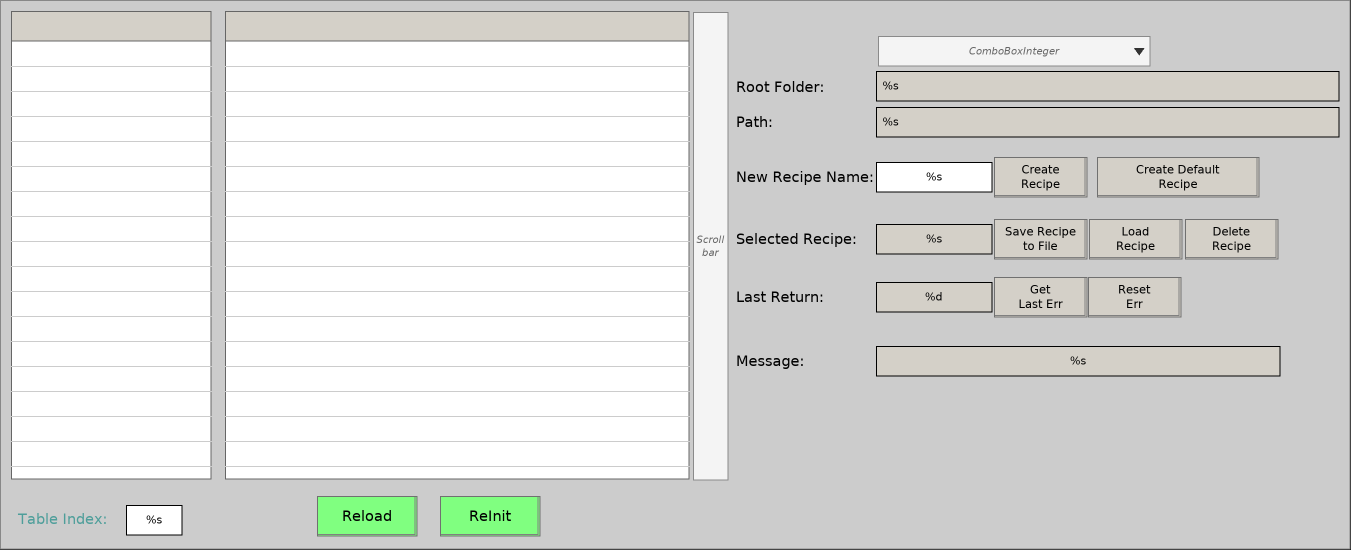
VISUALIZATION FB_Recipe_Vizu  // 1351x550
VAR_IN_OUT
	fb_Recipe		:FB_Recipe;
END_VAR
    Rectangle (0,0 1351x550)
    Table (11,11 200x468), data array: fb_Recipe.pstRecipe^.arrRecipeNames
        p1137915858: fb_Recipe.pstRecipe^.iRecipeIndex
        p1822360349: fb_Recipe.pstRecipe^.bValidSelected
        p3854506369: fb_Recipe.pstRecipe^.arrRecipeNames[INDEX]
        p2232123230: Recipe Names
    Rectangle (126,505 56x30), "%s", text variable: fb_Recipe.pstRecipe^.iRecipeIndex
    Label (15,504 108x30), "Table Index:"
    Button (317,496 100x40), "Reload"
        toggle fb_Recipe.pstRecipe^.bReloadRecipes
    Table (225,11 464x468), data array: fb_Recipe.pstRecipe^.arrVariableDisp
        p3854506369: fb_Recipe.pstRecipe^.arrVariableDisp[0,INDEX]
        p2232123230: No
        p1892666644: fb_Recipe.pstRecipe^.arrVariableDisp[1,INDEX]
        p511219082: Variable Name
        p338671338: fb_Recipe.pstRecipe^.arrVariableDisp[2,INDEX]
        p1755163831: Variable Value
    Scrollbar (693,12 35x468)
        p1057716461: fb_Recipe.pstRecipe^.iDispSel
    Button (1185,219 93x40), "Delete Recipe"
        toggle fb_Recipe.pstRecipe^.bDeleteRecipe
    Label (733,162 141x30), "New Recipe Name:"
    Label (733,224 141x30), "Selected Recipe:"
    Label (733,282 141x30), "Last Return:"
    Rectangle (876,162 116x30), "%s", text variable: fb_Recipe.pstRecipe^.sNewRecipeName
        OnMouseClick: write the text variable via Edit
    Rectangle (876,224 116x30), "%s", text variable: fb_Recipe.pstRecipe^.sSelectedReceipe
    Rectangle (876,282 116x30), "%d", text variable: fb_Recipe.LastReturn, colour toggle: fb_Recipe.LastReturn<>0
    Button (994,157 93x40), "Create Recipe"
        toggle fb_Recipe.pstRecipe^.bCreateRecipe
    Button (994,219 93x40), "Save Recipe to File"
        toggle fb_Recipe.pstRecipe^.bSaveFileCmd
    Button (994,277 93x40), "Get Last Err"
        toggle fb_Recipe.pstRecipe^.bGetLastError
    Button (1089,219 93x40), "Load Recipe"
        toggle fb_Recipe.pstRecipe^.bWriteToPLC_Cmd
    Button (1088,277 93x40), "Reset Err"
        toggle fb_Recipe.pstRecipe^.bResetLastError
    Label (733,107 141x30), "Path:"
    Rectangle (876,107 463x30), "%s", text variable: fb_Recipe.sRecipesStoragePath
    Button (440,496 100x40), "ReInit"
        toggle fb_Recipe.pstRecipe^.bReInit
    Label (733,346 141x30), "Message:"
    Rectangle (876,346 404x30), "%s", text variable: fb_Recipe.sMessage
    Button (1097,157 162x40), "Create Default Recipe"
        toggle fb_Recipe.pstRecipe^.bCreateRecipe
        OnMouseClick: execute { fb_Recipe.pstRecipe^.sNewRecipeName:='Default'; }
    ComboBoxInteger (878,36 272x30), variable: GVL_Recipe.eRecipeRootFolder, text list: 'TextList_RecipeRootFolder'
    Rectangle (876,71 463x30), "%s", text variable: GVL_Recipe.ar_RecipesStoragePath_Root[GVL_Recipe.eRecipeRootFolder]
        OnMouseClick: write the text variable via Edit
    Label (733,72 141x30), "Root Folder:"
END_VISUALIZATION

(* stored: Version 1.1.0.1, ProductVersion 3.1.4024.12
   Visu FB_Recipe_Vizu: Id {7547d88a-e051-4b2b-8116-5645fccffffe} *)
